Fanuc KAREL source: KT00857.KL

PROGRAM KT00857
%NOLOCKGROUP
VAR
  I1: INTEGER
  I2: INTEGER
  OUT: REAL
BEGIN
  I1 = 2
  I2 = 3
  I1 = 2
  I2 = 3
  OUT = ROUND(I1)
END KT00857
